ABB RAPID module: EdgeProg.mod

%%%
  VERSION:1
  LANGUAGE:ENGLISH
%%%
MODULE MOD_EdgeProg

    ! -------------------------------
    ! Define customized variables here
    ! ...

	! Tool variables:
	PERS tooldata ToolEdge := [TRUE,[[-1.500,2.250,99.875],[0.27059805,-0.65328148,0.65328148,0.27059805]],[1,[0,0,20],[1,0,0,0],0,0,0.005]];

	! Reference variables:
	PERS wobjdata FrameEdge := [FALSE, TRUE, "", [[0,0,0],[1,0,0,0]],[[100.500,-200.250,300.125],[0.94371436,0.26853582,-0.14487813,0.12767944]]];

	PROC Main()
		ConfJ \On;
		ConfL \Off;
		! Program generated by RoboDK v6.0.7 for ABB IRB 260 on XX/XX/XXXX 18:00:00
		! Using nominal kinematics.
		MoveAbsJ [[-15.000000,40.000000,20.000000,90.000000,0.000000,0.000000],[9E+09,9E+09,9E+09,9E+09,9E+09,9E+09]],[123.46,500,5000,1000],fine,ToolEdge \WObj:=FrameEdge;
		MoveL [[-624.230,571.208,454.620],[0.55239178,-0.04267608,0.67304167,-0.48995609],[0,0,0,1],[9E+09,9E+09,9E+09,9E+09,9E+09,9E+09]],[123.46,500,5000,1000],[FALSE,12.5,18.8,18.8,1.9,18.8,1.9],ToolEdge \WObj:=FrameEdge;
		STOP;
		WaitTime 1.234;
		TPWrite "A long message with "quotes", 'apostrophes' & symbols: <>[]{}()=+-*/%;#@! and more text to make it longer than eighty characters";
		! Comment with ; semicolon
		SetDO Gripper, ON;
		SetDO D_OUT_12, 0;
		SetAO Pressure, 0.75;
		WaitDI PartPresent, 1, \MaxTime:=0.2;
		WaitDI D_IN_7, 1;
		Do_Something 1, 2;
		x = 1
		MoveAbsJ [[30.000000,25.000000,80.000000,-45.000000,0.000000,0.000000],[9E+09,9E+09,9E+09,9E+09,9E+09,9E+09]],[123.46,500,5000,1000],[FALSE,12.5,18.8,18.8,1.9,18.8,1.9],ToolEdge \WObj:=FrameEdge;
	ENDPROC

ENDMODULE
